(* IEC 61131-3 sources: trust-platform/examples/OSCAT/pharma_filling_builder_state/oop/src, 3 files *)

(* ---- Main.st ---- *)
(* Record role: FillRecipe is a deterministic PLC-side record for tests and runtime readers. *)
TYPE FillRecipe :
STRUCT
    VolumeMl : REAL;
    PumpSpeedPct : REAL;
    LowWeightG : REAL;
    HighWeightG : REAL;
    Valid : BOOL;
END_STRUCT
END_TYPE

(* Composition role: FillRecipeBuilder owns the collaborating objects used by this Builder and State example. *)
FUNCTION_BLOCK FillRecipeBuilder
VAR
    Recipe : FillRecipe;
END_VAR

METHOD PUBLIC Reset
Recipe.VolumeMl := REAL#0.0;
Recipe.PumpSpeedPct := REAL#0.0;
Recipe.LowWeightG := REAL#0.0;
Recipe.HighWeightG := REAL#0.0;
Recipe.Valid := FALSE;
END_METHOD

METHOD PUBLIC SetVolume : FillRecipeBuilder
VAR_INPUT
    VolumeMl : REAL;
END_VAR
Recipe.VolumeMl := VolumeMl;
SetVolume := THIS;
END_METHOD

METHOD PUBLIC SetPumpSpeed : FillRecipeBuilder
VAR_INPUT
    PumpSpeedPct : REAL;
END_VAR
Recipe.PumpSpeedPct := PumpSpeedPct;
SetPumpSpeed := THIS;
END_METHOD

METHOD PUBLIC SetWeightWindow : FillRecipeBuilder
VAR_INPUT
    LowWeightG : REAL;
    HighWeightG : REAL;
END_VAR
Recipe.LowWeightG := LowWeightG;
Recipe.HighWeightG := HighWeightG;
SetWeightWindow := THIS;
END_METHOD

METHOD PUBLIC Build : FillRecipe
Recipe.Valid := (Recipe.VolumeMl > REAL#0.0) AND (Recipe.VolumeMl <= REAL#100.0) AND (Recipe.PumpSpeedPct > REAL#0.0) AND (Recipe.PumpSpeedPct <= REAL#100.0) AND (Recipe.HighWeightG > Recipe.LowWeightG);
Build := Recipe;
END_METHOD
END_FUNCTION_BLOCK

(* Pattern role: IFillingState is the contract boundary for the Builder and State example. *)
INTERFACE IFillingState
    PROPERTY StateId : INT
    GET
    END_GET
    END_PROPERTY

    METHOD OnExecute : INT
    VAR_INPUT
        StartCommand : BOOL;
        VialPresent : BOOL;
        FillDone : BOOL;
        WeightG : REAL;
        Recipe : FillRecipe;
    END_VAR
    END_METHOD
END_INTERFACE

(* Pattern role: IdleFillState is a concrete implementation in the Builder and State example. *)
FUNCTION_BLOCK IdleFillState IMPLEMENTS IFillingState
METHOD PUBLIC OnExecute : INT
VAR_INPUT
    StartCommand : BOOL;
    VialPresent : BOOL;
    FillDone : BOOL;
    WeightG : REAL;
    Recipe : FillRecipe;
END_VAR
IF StartCommand AND VialPresent AND Recipe.Valid THEN
    OnExecute := INT#10;
ELSE
    OnExecute := INT#0;
END_IF;
END_METHOD

PUBLIC PROPERTY StateId : INT
GET
    StateId := INT#0;
END_GET
END_PROPERTY
END_FUNCTION_BLOCK

(* Pattern role: PrimeFillState is a concrete implementation in the Builder and State example. *)
FUNCTION_BLOCK PrimeFillState IMPLEMENTS IFillingState
METHOD PUBLIC OnExecute : INT
VAR_INPUT
    StartCommand : BOOL;
    VialPresent : BOOL;
    FillDone : BOOL;
    WeightG : REAL;
    Recipe : FillRecipe;
END_VAR
OnExecute := INT#20;
END_METHOD

PUBLIC PROPERTY StateId : INT
GET
    StateId := INT#10;
END_GET
END_PROPERTY
END_FUNCTION_BLOCK

(* Pattern role: FillState is a concrete implementation in the Builder and State example. *)
FUNCTION_BLOCK FillState IMPLEMENTS IFillingState
METHOD PUBLIC OnExecute : INT
VAR_INPUT
    StartCommand : BOOL;
    VialPresent : BOOL;
    FillDone : BOOL;
    WeightG : REAL;
    Recipe : FillRecipe;
END_VAR
IF FillDone THEN
    OnExecute := INT#30;
ELSE
    OnExecute := INT#20;
END_IF;
END_METHOD

PUBLIC PROPERTY StateId : INT
GET
    StateId := INT#20;
END_GET
END_PROPERTY
END_FUNCTION_BLOCK

(* Pattern role: CheckWeightState is a concrete implementation in the Builder and State example. *)
FUNCTION_BLOCK CheckWeightState IMPLEMENTS IFillingState
METHOD PUBLIC OnExecute : INT
VAR_INPUT
    StartCommand : BOOL;
    VialPresent : BOOL;
    FillDone : BOOL;
    WeightG : REAL;
    Recipe : FillRecipe;
END_VAR
IF (WeightG >= Recipe.LowWeightG) AND (WeightG <= Recipe.HighWeightG) THEN
    OnExecute := INT#100;
ELSE
    OnExecute := INT#40;
END_IF;
END_METHOD

PUBLIC PROPERTY StateId : INT
GET
    StateId := INT#30;
END_GET
END_PROPERTY
END_FUNCTION_BLOCK

(* Pattern role: RejectState is a concrete implementation in the Builder and State example. *)
FUNCTION_BLOCK RejectState IMPLEMENTS IFillingState
METHOD PUBLIC OnExecute : INT
VAR_INPUT
    StartCommand : BOOL;
    VialPresent : BOOL;
    FillDone : BOOL;
    WeightG : REAL;
    Recipe : FillRecipe;
END_VAR
(* Restart-friendly terminal state: if a new vial is started in the
   same scan, jump to Prime so the next vial doesn't lose the start
   pulse waiting in Idle. *)
IF StartCommand AND VialPresent AND Recipe.Valid THEN
    OnExecute := INT#10;
ELSE
    OnExecute := INT#0;
END_IF;
END_METHOD

PUBLIC PROPERTY StateId : INT
GET
    StateId := INT#40;
END_GET
END_PROPERTY
END_FUNCTION_BLOCK

(* Pattern role: CompleteState is a concrete implementation in the Builder and State example. *)
FUNCTION_BLOCK CompleteState IMPLEMENTS IFillingState
METHOD PUBLIC OnExecute : INT
VAR_INPUT
    StartCommand : BOOL;
    VialPresent : BOOL;
    FillDone : BOOL;
    WeightG : REAL;
    Recipe : FillRecipe;
END_VAR
(* Same restart-friendly behavior as Reject: a fresh start pulse
   advances directly to Prime without going through Idle first. *)
IF StartCommand AND VialPresent AND Recipe.Valid THEN
    OnExecute := INT#10;
ELSE
    OnExecute := INT#0;
END_IF;
END_METHOD

PUBLIC PROPERTY StateId : INT
GET
    StateId := INT#100;
END_GET
END_PROPERTY
END_FUNCTION_BLOCK

(* Pattern role: FaultFillState is a concrete implementation in the Builder and State example. *)
FUNCTION_BLOCK FaultFillState IMPLEMENTS IFillingState
METHOD PUBLIC OnExecute : INT
VAR_INPUT
    StartCommand : BOOL;
    VialPresent : BOOL;
    FillDone : BOOL;
    WeightG : REAL;
    Recipe : FillRecipe;
END_VAR
OnExecute := INT#90;
END_METHOD

PUBLIC PROPERTY StateId : INT
GET
    StateId := INT#90;
END_GET
END_PROPERTY
END_FUNCTION_BLOCK

(* Composition role: FillingController owns the collaborating objects used by this Builder and State example. *)
FUNCTION_BLOCK FillingController
VAR
    Idle : IdleFillState;
    Prime : PrimeFillState;
    Filling : FillState;
    CheckWeight : CheckWeightState;
    Reject : RejectState;
    Complete : CompleteState;
    Fault : FaultFillState;
    Current : IFillingState;
    CurrentStateIdValue : INT;
    RejectCounter : DwordCounter;
    RecipeValue : FillRecipe;
END_VAR

METHOD PUBLIC Initialize
Current := Idle;
CurrentStateIdValue := INT#0;
RejectCounter.Initialize();
RejectCounter.Configure(StepSize := DWORD#1, MaxValue := DWORD#16#FFFFFFFF);
END_METHOD

METHOD PUBLIC LoadRecipe
VAR_INPUT
    Recipe : FillRecipe;
END_VAR
RecipeValue := Recipe;
END_METHOD

METHOD PUBLIC ResolveState : IFillingState
VAR_INPUT
    NextId : INT;
END_VAR
IF NextId = INT#10 THEN
    ResolveState := Prime;
ELSIF NextId = INT#20 THEN
    ResolveState := Filling;
ELSIF NextId = INT#30 THEN
    ResolveState := CheckWeight;
ELSIF NextId = INT#40 THEN
    ResolveState := Reject;
ELSIF NextId = INT#100 THEN
    ResolveState := Complete;
ELSIF NextId = INT#90 THEN
    ResolveState := Fault;
ELSE
    ResolveState := Idle;
END_IF;
END_METHOD

METHOD PUBLIC Update : INT
VAR_INPUT
    StartCommand : BOOL;
    VialPresent : BOOL;
    FillDone : BOOL;
    WeightG : REAL;
END_VAR
VAR
    NextId : INT;
END_VAR
NextId := Current.OnExecute(StartCommand := StartCommand, VialPresent := VialPresent, FillDone := FillDone, WeightG := WeightG, Recipe := RecipeValue);
IF NextId <> CurrentStateIdValue THEN
    Current := ResolveState(NextId := NextId);
    CurrentStateIdValue := NextId;
    IF NextId = INT#40 THEN
        (* COUNT_DR is edge-triggered; drop UP edge first so consecutive
           rejects across vials each register a fresh rising edge. *)
        RejectCounter.Update(Up := FALSE, Down := FALSE);
        RejectCounter.Update(Up := TRUE, Down := FALSE);
    END_IF;
END_IF;
Update := CurrentStateIdValue;
END_METHOD

PUBLIC PROPERTY CurrentStateId : INT
GET
    CurrentStateId := CurrentStateIdValue;
END_GET
END_PROPERTY

PUBLIC PROPERTY RejectCount : DWORD
GET
    RejectCount := RejectCounter.Count;
END_GET
END_PROPERTY

PUBLIC PROPERTY RecipeValid : BOOL
GET
    RecipeValid := RecipeValue.Valid;
END_GET
END_PROPERTY
END_FUNCTION_BLOCK

(* Scan role: Main wires the example objects and exposes the PLC call path under test. *)
PROGRAM Main
VAR
    Builder : FillRecipeBuilder;
    Filler : FillingController;
    StartCommand : BOOL;
    VialPresent : BOOL;
    FillDone : BOOL;
    WeightRaw : INT;
    Recipe : FillRecipe;
    PumpRunOut : BOOL;
    RejectOut : BOOL;
END_VAR

Recipe := Builder.SetVolume(VolumeMl := REAL#10.0).SetPumpSpeed(PumpSpeedPct := REAL#45.0).SetWeightWindow(LowWeightG := REAL#9.8, HighWeightG := REAL#10.2).Build();
Filler.Initialize();
Filler.LoadRecipe(Recipe := Recipe);
Filler.Update(StartCommand := StartCommand, VialPresent := VialPresent, FillDone := FillDone, WeightG := INT_TO_REAL(WeightRaw) / REAL#10.0);
PumpRunOut := Filler.CurrentStateId = INT#20;
RejectOut := Filler.CurrentStateId = INT#40;
END_PROGRAM

(* ---- Configuration.st ---- *)
CONFIGURATION PharmaFillingBuilderStateOopConfiguration
RESOURCE PharmaFillingBuilderStateOop ON PLC
    TASK MainTask (INTERVAL := T#50ms, PRIORITY := 1);
    PROGRAM Filler WITH MainTask : Main;
END_RESOURCE
VAR_CONFIG
    Filler.StartCommand AT %IX0.0 : BOOL;
    Filler.VialPresent AT %IX0.1 : BOOL;
    Filler.FillDone AT %IX0.2 : BOOL;
    Filler.WeightRaw AT %IW2 : INT;
    Filler.PumpRunOut AT %QX0.0 : BOOL;
    Filler.RejectOut AT %QX0.1 : BOOL;
END_VAR
END_CONFIGURATION

(* ---- Tests.st ---- *)
TEST_PROGRAM FillRecipeBuilderRejectsInvalidRecipe
VAR
    Builder : FillRecipeBuilder;
    Recipe : FillRecipe;
END_VAR

Recipe := Builder.SetVolume(VolumeMl := REAL#0.0).SetPumpSpeed(PumpSpeedPct := REAL#50.0).SetWeightWindow(LowWeightG := REAL#9.8, HighWeightG := REAL#10.2).Build();
ASSERT_FALSE(IN := Recipe.Valid);
END_TEST_PROGRAM

TEST_PROGRAM FillingStateObjectsRejectBadWeight
VAR
    Builder : FillRecipeBuilder;
    Recipe : FillRecipe;
    Filler : FillingController;
END_VAR

Recipe := Builder.SetVolume(VolumeMl := REAL#10.0).SetPumpSpeed(PumpSpeedPct := REAL#45.0).SetWeightWindow(LowWeightG := REAL#9.8, HighWeightG := REAL#10.2).Build();
Filler.Initialize();
Filler.LoadRecipe(Recipe := Recipe);
ASSERT_EQUAL(EXPECTED := INT#10, ACTUAL := Filler.Update(StartCommand := TRUE, VialPresent := TRUE, FillDone := FALSE, WeightG := REAL#0.0));
ASSERT_EQUAL(EXPECTED := INT#20, ACTUAL := Filler.Update(StartCommand := FALSE, VialPresent := TRUE, FillDone := FALSE, WeightG := REAL#0.0));
ASSERT_EQUAL(EXPECTED := INT#30, ACTUAL := Filler.Update(StartCommand := FALSE, VialPresent := TRUE, FillDone := TRUE, WeightG := REAL#0.0));
ASSERT_EQUAL(EXPECTED := INT#40, ACTUAL := Filler.Update(StartCommand := FALSE, VialPresent := TRUE, FillDone := FALSE, WeightG := REAL#10.5));
ASSERT_EQUAL(EXPECTED := DWORD#1, ACTUAL := Filler.RejectCount);
END_TEST_PROGRAM

(* Two-vial sequence test: drives one Filler through two complete
   fill cycles (one good, one bad). Catches bugs where reject counts
   leak between vials or where the state machine sticks at Reject
   after the first bad vial. *)
TEST_PROGRAM FillerProcessesMultipleVialsOnOneInstance
VAR
    Builder : FillRecipeBuilder;
    Recipe : FillRecipe;
    Filler : FillingController;
END_VAR

Recipe := Builder.SetVolume(VolumeMl := REAL#10.0).SetPumpSpeed(PumpSpeedPct := REAL#45.0).SetWeightWindow(LowWeightG := REAL#9.8, HighWeightG := REAL#10.2).Build();
Filler.Initialize();
Filler.LoadRecipe(Recipe := Recipe);

(* Vial 1: in-window weight (10.0 g) - should not increment reject *)
Filler.Update(StartCommand := TRUE, VialPresent := TRUE, FillDone := FALSE, WeightG := REAL#0.0);
Filler.Update(StartCommand := FALSE, VialPresent := TRUE, FillDone := FALSE, WeightG := REAL#0.0);
Filler.Update(StartCommand := FALSE, VialPresent := TRUE, FillDone := TRUE, WeightG := REAL#0.0);
Filler.Update(StartCommand := FALSE, VialPresent := TRUE, FillDone := FALSE, WeightG := REAL#10.0);
ASSERT_EQUAL(EXPECTED := DWORD#0, ACTUAL := Filler.RejectCount);

(* Vial 2: out-of-window weight (11 g) - reject increments *)
Filler.Update(StartCommand := TRUE, VialPresent := TRUE, FillDone := FALSE, WeightG := REAL#0.0);
Filler.Update(StartCommand := FALSE, VialPresent := TRUE, FillDone := FALSE, WeightG := REAL#0.0);
Filler.Update(StartCommand := FALSE, VialPresent := TRUE, FillDone := TRUE, WeightG := REAL#0.0);
Filler.Update(StartCommand := FALSE, VialPresent := TRUE, FillDone := FALSE, WeightG := REAL#11.0);
ASSERT_EQUAL(EXPECTED := DWORD#1, ACTUAL := Filler.RejectCount);
END_TEST_PROGRAM

(* Builder boundary tests: each validation rule trips correctly.
   Volume must be in (0, 100], pump speed in (0, 100], window
   non-empty (High > Low). *)
TEST_PROGRAM FillRecipeBuilderBoundaryValidation
VAR
    Builder : FillRecipeBuilder;
    Recipe : FillRecipe;
END_VAR

(* Volume too high - invalid *)
Builder.Reset();
Recipe := Builder.SetVolume(VolumeMl := REAL#150.0).SetPumpSpeed(PumpSpeedPct := REAL#50.0).SetWeightWindow(LowWeightG := REAL#9.8, HighWeightG := REAL#10.2).Build();
ASSERT_FALSE(IN := Recipe.Valid);

(* Pump speed too high - invalid *)
Builder.Reset();
Recipe := Builder.SetVolume(VolumeMl := REAL#10.0).SetPumpSpeed(PumpSpeedPct := REAL#120.0).SetWeightWindow(LowWeightG := REAL#9.8, HighWeightG := REAL#10.2).Build();
ASSERT_FALSE(IN := Recipe.Valid);

(* Weight window inverted - invalid *)
Builder.Reset();
Recipe := Builder.SetVolume(VolumeMl := REAL#10.0).SetPumpSpeed(PumpSpeedPct := REAL#50.0).SetWeightWindow(LowWeightG := REAL#10.2, HighWeightG := REAL#9.8).Build();
ASSERT_FALSE(IN := Recipe.Valid);

(* Boundary upper edges: VolumeMl = 100, PumpSpeedPct = 100 are valid *)
Builder.Reset();
Recipe := Builder.SetVolume(VolumeMl := REAL#100.0).SetPumpSpeed(PumpSpeedPct := REAL#100.0).SetWeightWindow(LowWeightG := REAL#99.0, HighWeightG := REAL#101.0).Build();
ASSERT_TRUE(IN := Recipe.Valid);

(* Boundary zero: pump speed = 0 is invalid *)
Builder.Reset();
Recipe := Builder.SetVolume(VolumeMl := REAL#10.0).SetPumpSpeed(PumpSpeedPct := REAL#0.0).SetWeightWindow(LowWeightG := REAL#9.8, HighWeightG := REAL#10.2).Build();
ASSERT_FALSE(IN := Recipe.Valid);
END_TEST_PROGRAM

(* Recipe gating: Filler must refuse to leave Idle when the loaded
   recipe is invalid, regardless of StartCommand or VialPresent. *)
TEST_PROGRAM FillerHoldsAtIdleWhenRecipeInvalid
VAR
    Builder : FillRecipeBuilder;
    Recipe : FillRecipe;
    Filler : FillingController;
END_VAR

(* Build an invalid recipe (volume = 0) *)
Recipe := Builder.SetVolume(VolumeMl := REAL#0.0).SetPumpSpeed(PumpSpeedPct := REAL#45.0).SetWeightWindow(LowWeightG := REAL#9.8, HighWeightG := REAL#10.2).Build();
Filler.Initialize();
Filler.LoadRecipe(Recipe := Recipe);
ASSERT_FALSE(IN := Filler.RecipeValid);

(* All inputs healthy but recipe invalid: must hold at Idle *)
ASSERT_EQUAL(EXPECTED := INT#0, ACTUAL := Filler.Update(StartCommand := TRUE, VialPresent := TRUE, FillDone := FALSE, WeightG := REAL#0.0));
ASSERT_EQUAL(EXPECTED := INT#0, ACTUAL := Filler.Update(StartCommand := TRUE, VialPresent := TRUE, FillDone := TRUE, WeightG := REAL#10.0));

(* Reload with a valid recipe: now starts on next StartCommand *)
Recipe := Builder.SetVolume(VolumeMl := REAL#10.0).SetPumpSpeed(PumpSpeedPct := REAL#45.0).SetWeightWindow(LowWeightG := REAL#9.8, HighWeightG := REAL#10.2).Build();
Filler.LoadRecipe(Recipe := Recipe);
ASSERT_TRUE(IN := Filler.RecipeValid);
ASSERT_EQUAL(EXPECTED := INT#10, ACTUAL := Filler.Update(StartCommand := TRUE, VialPresent := TRUE, FillDone := FALSE, WeightG := REAL#0.0));
END_TEST_PROGRAM

(* Per-state isolation: each state FB returns its own id and computes
   transitions independent of any controller state. The state objects
   are not stateful - they read inputs and Recipe each call. *)
TEST_PROGRAM FillingStatesAreStatelessOracles
VAR
    Idle : IdleFillState;
    Prime : PrimeFillState;
    Fill : FillState;
    CheckWeight : CheckWeightState;
    Reject : RejectState;
    Complete : CompleteState;
    Recipe : FillRecipe;
END_VAR

(* StateId reflects the state's own number *)
ASSERT_EQUAL(EXPECTED := INT#0, ACTUAL := Idle.StateId);
ASSERT_EQUAL(EXPECTED := INT#10, ACTUAL := Prime.StateId);
ASSERT_EQUAL(EXPECTED := INT#20, ACTUAL := Fill.StateId);
ASSERT_EQUAL(EXPECTED := INT#30, ACTUAL := CheckWeight.StateId);
ASSERT_EQUAL(EXPECTED := INT#40, ACTUAL := Reject.StateId);
ASSERT_EQUAL(EXPECTED := INT#100, ACTUAL := Complete.StateId);

(* Make a valid recipe *)
Recipe.VolumeMl := REAL#10.0;
Recipe.PumpSpeedPct := REAL#45.0;
Recipe.LowWeightG := REAL#9.8;
Recipe.HighWeightG := REAL#10.2;
Recipe.Valid := TRUE;

(* Idle: with start + vial + valid recipe, advances to Prime *)
ASSERT_EQUAL(EXPECTED := INT#10, ACTUAL := Idle.OnExecute(StartCommand := TRUE, VialPresent := TRUE, FillDone := FALSE, WeightG := REAL#0.0, Recipe := Recipe));
(* Prime: always advances to Fill *)
ASSERT_EQUAL(EXPECTED := INT#20, ACTUAL := Prime.OnExecute(StartCommand := FALSE, VialPresent := TRUE, FillDone := FALSE, WeightG := REAL#0.0, Recipe := Recipe));
(* Fill: stays on no FillDone, advances on FillDone *)
ASSERT_EQUAL(EXPECTED := INT#20, ACTUAL := Fill.OnExecute(StartCommand := FALSE, VialPresent := TRUE, FillDone := FALSE, WeightG := REAL#0.0, Recipe := Recipe));
ASSERT_EQUAL(EXPECTED := INT#30, ACTUAL := Fill.OnExecute(StartCommand := FALSE, VialPresent := TRUE, FillDone := TRUE, WeightG := REAL#0.0, Recipe := Recipe));
(* CheckWeight: in window -> Complete; out of window -> Reject *)
ASSERT_EQUAL(EXPECTED := INT#100, ACTUAL := CheckWeight.OnExecute(StartCommand := FALSE, VialPresent := TRUE, FillDone := FALSE, WeightG := REAL#10.0, Recipe := Recipe));
ASSERT_EQUAL(EXPECTED := INT#40, ACTUAL := CheckWeight.OnExecute(StartCommand := FALSE, VialPresent := TRUE, FillDone := FALSE, WeightG := REAL#11.0, Recipe := Recipe));

(* Reject and Complete are restart-friendly: a fresh start advances to Prime *)
ASSERT_EQUAL(EXPECTED := INT#10, ACTUAL := Reject.OnExecute(StartCommand := TRUE, VialPresent := TRUE, FillDone := FALSE, WeightG := REAL#0.0, Recipe := Recipe));
ASSERT_EQUAL(EXPECTED := INT#10, ACTUAL := Complete.OnExecute(StartCommand := TRUE, VialPresent := TRUE, FillDone := FALSE, WeightG := REAL#0.0, Recipe := Recipe));
(* Without start: both return to Idle *)
ASSERT_EQUAL(EXPECTED := INT#0, ACTUAL := Reject.OnExecute(StartCommand := FALSE, VialPresent := TRUE, FillDone := FALSE, WeightG := REAL#0.0, Recipe := Recipe));
ASSERT_EQUAL(EXPECTED := INT#0, ACTUAL := Complete.OnExecute(StartCommand := FALSE, VialPresent := TRUE, FillDone := FALSE, WeightG := REAL#0.0, Recipe := Recipe));
END_TEST_PROGRAM

(* Builder reuse: after Build, calling Reset gives a fresh recipe
   without leaking the previous values. *)
TEST_PROGRAM FillRecipeBuilderResetClearsState
VAR
    Builder : FillRecipeBuilder;
    Recipe1 : FillRecipe;
    Recipe2 : FillRecipe;
END_VAR

Recipe1 := Builder.SetVolume(VolumeMl := REAL#10.0).SetPumpSpeed(PumpSpeedPct := REAL#45.0).SetWeightWindow(LowWeightG := REAL#9.8, HighWeightG := REAL#10.2).Build();
ASSERT_TRUE(IN := Recipe1.Valid);

(* Reset wipes the internal recipe; Build without setters yields
   invalid (volume = 0, pump = 0) *)
Builder.Reset();
Recipe2 := Builder.Build();
ASSERT_FALSE(IN := Recipe2.Valid);
ASSERT_NEAR(EXPECTED := REAL#0.0, ACTUAL := Recipe2.VolumeMl, DELTA := REAL#0.001);
ASSERT_NEAR(EXPECTED := REAL#0.0, ACTUAL := Recipe2.PumpSpeedPct, DELTA := REAL#0.001);

(* Original recipe1 is unchanged - the builder returned a copy *)
ASSERT_TRUE(IN := Recipe1.Valid);
ASSERT_NEAR(EXPECTED := REAL#10.0, ACTUAL := Recipe1.VolumeMl, DELTA := REAL#0.001);
END_TEST_PROGRAM
